(* IEC 61131-3 sources: llm-plc-st-eval/data/definitivo/qwen2.5-coder_14b/B2/few_shot, 3 files *)

(* ---- ejec_1.st ---- *)
FUNCTION_BLOCK FB_Valvula
VAR_INPUT
    nivelAlto : BOOL; (* Sensor de nivel alto *)
END_VAR
VAR_OUTPUT
    valvula : BOOL; (* Válvula de drenaje *)
END_VAR
VAR
    tNivelAlto : TP; (* Temporizador para el nivel alto *)
END_VAR

(* Temporiza el tiempo que el nivel está alto *)
tNivelAlto(IN := nivelAlto, PT := T#5S);

(* La válvula se abre si el nivel está alto durante 5 segundos *)
valvula := tNivelAlto.Q;

(* La válvula se cierra inmediatamente si el nivel deja de estar alto *)
IF NOT nivelAlto THEN
    valvula := FALSE;
END_IF
END_FUNCTION_BLOCK

(* ---- ejec_2.st ---- *)
FUNCTION_BLOCK FB_Valvula
VAR_INPUT
    nivelAlto : BOOL; (* Sensor de nivel alto *)
END_VAR
VAR_OUTPUT
    valvula : BOOL; (* Válvula de drenaje *)
END_VAR
VAR
    tNivelAlto : TP; (* Temporizador para el nivel alto *)
END_VAR

(* Temporizador que se activa cuando el nivel está alto *)
tNivelAlto(IN := nivelAlto, PT := T#5S);

(* La válvula se abre si el temporizador ha expirado *)
valvula := tNivelAlto.Q;

(* La válvula se cierra inmediatamente si el nivel deja de estar alto *)
IF NOT nivelAlto THEN
    valvula := FALSE;
END_IF
END_FUNCTION_BLOCK

(* ---- ejec_3.st ---- *)
FUNCTION_BLOCK FB_Valvula
VAR_INPUT
    nivelAlto : BOOL; (* Sensor de nivel alto *)
END_VAR
VAR_OUTPUT
    valvula : BOOL; (* Válvula de drenaje *)
END_VAR
VAR
    tNivel : TP; (* Temporizador para el nivel alto *)
END_VAR

(* Temporizador que se activa cuando el nivel está alto *)
tNivel(IN := nivelAlto, PT := T#5S);

(* La válvula se abre si el temporizador ha expirado *)
valvula := tNivel.Q;

(* La válvula se cierra inmediatamente si el nivel deja de estar alto *)
IF NOT nivelAlto THEN
    valvula := FALSE;
END_IF
END_FUNCTION_BLOCK
